FUNCTION_BLOCK "FB_PressDemoLoadPosition"
{ S7_Optimized_Access := 'TRUE' }
VERSION : 0.1
VAR_INPUT
    Run : Bool;
    Reset : Bool;
    OwnerIndex : DInt;
    ChainIndex : DInt;
    Delta : Time;
END_VAR
VAR_IN_OUT
    PressRam {ExternalAccessible := 'False'; ExternalVisible := 'False'; ExternalWritable := 'False'} : "FB_CylinderCM";
    Door {ExternalAccessible := 'False'; ExternalVisible := 'False'; ExternalWritable := 'False'} : "FB_CylinderCM";
    PartSlide {ExternalAccessible := 'False'; ExternalVisible := 'False'; ExternalWritable := 'False'} : "FB_CylinderCM";
END_VAR
VAR_OUTPUT
END_VAR
VAR
    Seq {ExternalWritable := 'False'} : "FRK_SequenceCtx";
    Row1 {ExternalWritable := 'False'} : "FRK_SequenceRow";
    Row2 {ExternalWritable := 'False'} : "FRK_SequenceRow";
    Row3 {ExternalWritable := 'False'} : "FRK_SequenceRow";
    Row4 {ExternalWritable := 'False'} : "FRK_SequenceRow";
    At240 {ExternalAccessible := 'False'; ExternalVisible := 'False'; ExternalWritable := 'False'} : Bool;
    At260 {ExternalAccessible := 'False'; ExternalVisible := 'False'; ExternalWritable := 'False'} : Bool;
    At280 {ExternalAccessible := 'False'; ExternalVisible := 'False'; ExternalWritable := 'False'} : Bool;
    At300 {ExternalAccessible := 'False'; ExternalVisible := 'False'; ExternalWritable := 'False'} : Bool;
    Ready1 {ExternalAccessible := 'False'; ExternalVisible := 'False'; ExternalWritable := 'False'} : Bool;
    Ready2 {ExternalAccessible := 'False'; ExternalVisible := 'False'; ExternalWritable := 'False'} : Bool;
    Ready3 {ExternalAccessible := 'False'; ExternalVisible := 'False'; ExternalWritable := 'False'} : Bool;
    Ready4 {ExternalAccessible := 'False'; ExternalVisible := 'False'; ExternalWritable := 'False'} : Bool;
    Ready5 {ExternalAccessible := 'False'; ExternalVisible := 'False'; ExternalWritable := 'False'} : Bool;
    Advance {ExternalAccessible := 'False'; ExternalVisible := 'False'; ExternalWritable := 'False'} : Bool;
END_VAR
BEGIN
    "FRK_SeqBegin"(Run := #Run, Reset := #Reset, OwnerIndex := #OwnerIndex, ChainIndex := #ChainIndex, BranchIndex := 1, ViewOffset := 360, ViewDepth := 1, Delta := #Delta, Seq := #Seq);
    "FRK_SeqInitial"(Seq := #Seq, InitialStep := 240);
    "F_CylinderSequenceLease"(Seq := #Seq, Target := #PressRam);
    "F_CylinderSequenceLease"(Seq := #Seq, Target := #Door);
    "F_CylinderSequenceLease"(Seq := #Seq, Target := #PartSlide);
    CASE #Seq.ScanStep OF
        240:
            IF #Seq.Running AND NOT #Seq.Error THEN
                "FRK_SeqStep"(StepNo := 240, StepName := 'project.step.pressReturnRam', AwaitingLabel := 'PressRam.RETRACT', AwaitsPath := #PressRam.Status.Name, TimeClass := 0, ExpectedTime := #Seq.NoTimeGuard, Seq := #Seq, Row := #Row1);
                #Ready1 := "F_CylinderRetract"(Seq := #Seq, Target := #PressRam);
                "FRK_SeqReady"(Seq := #Seq, Ok1 := #Ready1, Ok2 := TRUE, Ok3 := TRUE, Ok4 := TRUE, Ok5 := TRUE);
                "FRK_SeqRoute"(Seq := #Seq, OnAdvance := 260, OnJump1 := -1);
            END_IF;
        260:
            IF #Seq.Running AND NOT #Seq.Error THEN
                "FRK_SeqStep"(StepNo := 260, StepName := 'project.step.pressReturnDoor', AwaitingLabel := 'Door.RETRACT', AwaitsPath := #Door.Status.Name, TimeClass := 0, ExpectedTime := #Seq.NoTimeGuard, Seq := #Seq, Row := #Row2);
                #Ready1 := "F_CylinderRetract"(Seq := #Seq, Target := #Door);
                "FRK_SeqReady"(Seq := #Seq, Ok1 := #Ready1, Ok2 := TRUE, Ok3 := TRUE, Ok4 := TRUE, Ok5 := TRUE);
                "FRK_SeqRoute"(Seq := #Seq, OnAdvance := 280, OnJump1 := -1);
            END_IF;
        280:
            IF #Seq.Running AND NOT #Seq.Error THEN
                "FRK_SeqStep"(StepNo := 280, StepName := 'project.step.pressReturnSlide', AwaitingLabel := 'PartSlide.RETRACT', AwaitsPath := #PartSlide.Status.Name, TimeClass := 0, ExpectedTime := #Seq.NoTimeGuard, Seq := #Seq, Row := #Row3);
                #Ready1 := "F_CylinderRetract"(Seq := #Seq, Target := #PartSlide);
                "FRK_SeqReady"(Seq := #Seq, Ok1 := #Ready1, Ok2 := TRUE, Ok3 := TRUE, Ok4 := TRUE, Ok5 := TRUE);
                "FRK_SeqRoute"(Seq := #Seq, OnAdvance := 300, OnJump1 := -1);
            END_IF;
        300:
            IF #Seq.Running AND NOT #Seq.Error THEN
                "FRK_SeqStep"(StepNo := 300, StepName := 'project.step.pressLoadPositionComplete', AwaitingLabel := '', AwaitsPath := '', TimeClass := 0, ExpectedTime := #Seq.NoTimeGuard, Seq := #Seq, Row := #Row4);
                "FRK_SeqComplete"(Seq := #Seq);
            END_IF;
        ELSE
            IF #Seq.Running AND NOT #Seq.Error THEN
                #Seq.Error := TRUE;
                #Seq.ErrorDiagnostic.ReasonCode := 10001;
                #Seq.ErrorDiagnostic.Description := WSTRING#'project.sequence.invalidStep';
            END_IF;
    END_CASE;
    "F_CylinderSequenceLease"(Seq := #Seq, Target := #PressRam);
    "F_CylinderSequenceLease"(Seq := #Seq, Target := #Door);
    "F_CylinderSequenceLease"(Seq := #Seq, Target := #PartSlide);
END_FUNCTION_BLOCK
FUNCTION "F_PressDemoLoadPosition" : Bool
{ S7_Optimized_Access := 'TRUE' }
VERSION : 0.1
VAR_INPUT Run : Bool; Reset : Bool; OwnerIndex : DInt; ChainIndex : DInt; Delta : Time; END_VAR
VAR_IN_OUT Target : "FB_PressDemoLoadPosition"; PressRam : "FB_CylinderCM"; Door : "FB_CylinderCM"; PartSlide : "FB_CylinderCM"; END_VAR
BEGIN
    // Each embedding chain passes its own identity, so two owners of the one
    // motion chain never share a command lease.
    #Target(Run := #Run, Reset := #Reset, OwnerIndex := #OwnerIndex, ChainIndex := #ChainIndex, Delta := #Delta, PressRam := #PressRam, Door := #Door, PartSlide := #PartSlide);
    #F_PressDemoLoadPosition := #Target.Seq.Done;
END_FUNCTION
